(* IEC 61131-3 sources: bevling_machine/framework/sources/00_Types, 16 files *)

(* ---- E_AutoStep.st ---- *)
(* 模块说明：自动主流程步骤。正常循环从送料等料开始，切割完成后执行三路收尾。 *)
{attribute 'qualified_only'}
TYPE E_AutoStep :
(
    Idle := 0, (* 主流程待机 *)
    FeedWait := 10, (* 正常送料等料，可长期等待 *)
    StopFeed := 20, (* 撤销皮带运行并等待停止 *)
    Push := 30, (* G3 推动气缸动作 *)
    Clearance := 40, (* 并行避让 P/Q，全完成后继续 *)
    Rotate := 50, (* D8 平台旋转到配方角度 *)
    PressDown := 60, (* G1 下压到位 *)
    KnifeDown := 70, (* G9 盘刀下降到位 *)
    SpindleOn := 80, (* D3 盘刀运行状态建立 *)
    Cutting := 90, (* D2 走刀和 G6 吹气，等待指定行程到位 *)
    StopCut := 100, (* 停止盘刀和吹气 *)
    PostCut := 110, (* 抬刀、抬压、并行三路收尾 *)
    Complete := 120, (* 整循环完成，连续模式回送料 *)
    Fault := 900 (* 自动流程错误，退出执行后复位 *)
);
END_TYPE

(* ---- E_DeviceAction.st ---- *)
(* 模块说明：统一设备动作类型。未请求或停止时取消动作；定位完成依据本次命令序号判断。 *)
{attribute 'qualified_only'}
TYPE E_DeviceAction :
(
    None := 0, (* 无动作请求，取消当前动作 *)
    Position := 1, (* 定位到指定目标，等待本次序号完成 *)
    Run := 2, (* 保持连续运行请求 *)
    Jog := 3, (* 保持点动，速度正负决定方向 *)
    Stop := 4, (* 取消动作，停止运行 *)
    Home := 5 (* 回零：按轴配置的回零方式寻找原点，完成后把轴坐标设为回零坐标 *)
);
END_TYPE

(* ---- E_DeviceKind.st ---- *)
(* 模块说明：设备适配类型，由设备管理器选择轴、电机、气缸或阀的执行入口。 *)
{attribute 'qualified_only'}
TYPE E_DeviceKind :
(
    Unused := 0, (* 保留，不调度 *)
    Axis := 1, (* 定位轴 *)
    Motor := 2, (* 连续电机 *)
    Cylinder := 3, (* 两端动作气缸 *)
    Valve := 4 (* 开关阀 *)
);
END_TYPE

(* ---- E_MachineMode.st ---- *)
(* 模块说明：操作模式。手动与自动分别提出动作请求，共用设备执行和互锁。 *)
{attribute 'qualified_only'}
TYPE E_MachineMode :
(
    Manual := 0, (* 手动点动/单机构调试 *)
    Automatic := 1 (* 自动循环工序 *)
);
END_TYPE

(* ---- E_MachineState.st ---- *)
(* 模块说明：整机运行状态。停止或报警复位后须重新初始化，启动命令不会跳过初始化。 *)
{attribute 'qualified_only'}
TYPE E_MachineState :
(
    Stopped := 0, (* 停止，须初始化 *)
    Initializing := 10, (* 初始化中 *)
    Ready := 20, (* 初始化完成，等待自动启动 *)
    Manual := 30, (* 手动控制中 *)
    Automatic := 40, (* 自动工序运行中，包含正常等料 *)
    Fault := 90 (* 报警锁存，清除原因后复位 *)
);
END_TYPE

(* ---- ST_DeviceCommand.st ---- *)
(* 模块说明：上层发给单个设备的请求。定位每次换新序号；连续运行和点动期间保持请求。 *)
TYPE ST_DeviceCommand :
STRUCT
eAction : E_DeviceAction; (* 动作类型：无请求、定位、连续运行、点动或停止，见 E_DeviceAction。 *)
udiID : UDINT; (* 本次命令序号，0 无效；发起新定位时换新序号。 *)
lrTarget : LREAL; (* 目标工程位置；气缸使用约定的 0/1 端点，连续运行和点动不使用该位置。 *)
lrVelocity : LREAL; (* 请求速度，单位随设备工程单位定义；尚未完成实机标定。 *)
END_STRUCT
END_TYPE

(* ---- ST_DeviceConfig.st ---- *)
(* 模块说明：设备类型、行程范围和仿真参数。当前工程单位与时间均为仿真示例，尚未完成实机标定。 *)
TYPE ST_DeviceConfig :
STRUCT
	eKind : E_DeviceKind; (* 设备类型，决定调用哪一种设备适配功能块。 *)
	lrInitialPosition : LREAL; (* 首次进入仿真时的初始位置，不是实机回原点结果。 *)
	lrMinPosition : LREAL := -1000.0; (* 示例软行程下限，单位随机构定义。 *)
	lrMaxPosition : LREAL := 1000.0; (* 示例软行程上限，单位随机构定义。 *)
	lrMaxVelocity : LREAL := 100.0; (* 允许请求的最大速度，用于仿真命令范围检查。 *)
	tSimAction : TIME := T#500MS; (* 仿真单次定位/建立运行状态所需时间，不代表实际机械动作时间。 *)
	lrMaxAcceleration : LREAL := 50.0; (* 真实轴加速度上限，mm/s2；仿真不使用该字段。 *)
	lrMaxDeceleration : LREAL := 50.0; (* 真实轴减速度上限，mm/s2；仿真不使用该字段。 *)
	xAbsoluteAllowed : BOOL := FALSE; (* 真实轴是否允许绝对定位；未回零时必须保持 FALSE。 *)
END_STRUCT
END_TYPE

(* ---- ST_DeviceStatus.st ---- *)
(* 模块说明：单个设备的执行反馈。收到命令与完成命令是两个状态，不能只看忙标志判断完成。 *)
TYPE ST_DeviceStatus :
STRUCT
xReady : BOOL; (* 设备已使能且无故障，允许接收命令；不表示动作已经完成。 *)
xBusy : BOOL; (* 当前动作正在执行，定位完成或停止后清除。 *)
xActive : BOOL; (* 连续运行已建立或点动正在进行；定位动作完成后不保持该标志。 *)
xError : BOOL; (* 本设备或本子流程发生故障；具体原因见对应错误码。 *)
udiErrorID : UDINT; (* 错误码；0 表示无错误，设备或流程发生异常时赋值。 *)
udiAcceptedID : UDINT; (* 设备已接收的命令序号，用于区别尚未接收与正在执行。 *)
udiCompletedID : UDINT; (* 设备已完成的命令序号；应与本次 udiID 匹配后再切换步骤。 *)
lrPosition : LREAL; (* 实际或仿真反馈位置；气缸 0/1 的方向见设备编号说明。 *)
xRealActive : BOOL; (* TRUE 表示该编号当前由真实执行后端接管，不是仿真模型；默认 FALSE。 *)
xHomed : BOOL; (* 真实轴本次上电后已完成回零；仿真设备恒为 FALSE。回零成功前绝对定位会被拒绝。 *)
END_STRUCT
END_TYPE

(* ---- ST_MachineStatus.st ---- *)
(* 模块说明：提供给监控和上位机的整机状态。可从主步骤、支线步骤、报警和互锁阻挡编号定位等待原因。 *)
TYPE ST_MachineStatus :
STRUCT
	eState : E_MachineState; (* 整机状态，见 E_MachineState；调试时先确认是否已初始化及处于正确模式。 *)
	eMode : E_MachineMode; (* 本地模式旋钮的当前选择：Manual 手动，Automatic 自动；上位机仅可读取。 *)
	eAutoStep : E_AutoStep; (* 自动主流程步骤；送料、避让、切割、收尾等状态见 E_AutoStep。 *)
	xSimulation : BOOL; (* TRUE 使用内部仿真；当前 FALSE 报未实现 3001，不会接管真实运动。 *)
	xRealBackendAvailable : BOOL; (* 真实设备适配是否已具备；当前框架固定 FALSE。 *)
	xRemoteStartStopAllowed : BOOL; (* 当前是否允许上位机启停，供只读状态发布；与物理手动/自动模式独立。 *)
	xInitialized : BOOL; (* 初始化完成标志；停止、运行中切换模式或故障会清除。 *)
	xReady : BOOL; (* 整机已经初始化并处于 Ready 状态，可接受自动启动；手动状态下不置该位。 *)
	xMaterialAtLength : BOOL; (* 定长光电到位状态；自动送料须先离开再到位，并满足 D5 下降。 *)
	xCycleComplete : BOOL; (* 一个扫描周期的整循环完成脉冲，可用于计数或上位机提示。 *)
	udiCycleCount : UDINT; (* 已完成的自动整循环计数；包括机械手移料等三路收尾。 *)
	udiAlarm : UDINT; (* 整机锁存报警码；0 无报警，1001 安全许可，3001 实机未接入，10000+索引为设备故障。 *)
	uiBlockedDevice : UINT; (* 本扫描最后一个被互锁阻挡的设备索引；0 表示无阻挡，可结合设备状态排查。 *)
	uiManualReject : UINT; (* 本扫描最后一个被拒绝的手动设备索引；0 无拒绝，检查相反按钮或动作类型。 *)
	uiClearLengthStep : UINT; (* 避让支线 P 的当前步骤：10 升起 D5，20 移开 D4，1000 完成。 *)
	uiClearTransferStep : UINT; (* 避让支线 Q 当前步骤：10 降 G4，20 松 G3，30 降 G2，1000 完成。 *)
	uiPostStep : UINT; (* 收尾总步骤：10 抬刀，20 抬压，30 等待三路完成，1000 结束。 *)
	uiReturnKnifeStep : UINT; (* 收尾支线 A：10 喷油，20 D2 回刀，1000 完成。 *)
	uiUnloadStep : UINT; (* 机械手移料支线 B 步骤，10..110 每步加 10，1000 完成；详见 FB_Unload。 *)
	uiResetLengthStep : UINT; (* 收尾支线 C：10 D4 定位，20 D5 下降，30 确认下降，1000 完成。 *)
	uiInitializeStep : UINT; (* 初始化步骤：10 整理刀/压/夹爪，20 避让，25 真实轴回零，30 初始定位，40 定长下降，1000 完成。 *)
	uiActiveMaterialModel : UINT; (* 已采纳的运行料型，取自运行配方；可能与尚未生效的参数区不同。 *)
	wRemoteAckSequence : WORD; (* 整机已处理的上位机命令序号；应结合 uiRemoteResult 判断是否接受。 *)
	uiRemoteResult : UINT; (* 远程处理结果：0 接受，1 未授权，2 不支持命令，3 状态/本地停止不允许，4 验证模式禁止自动，5 配方不合法。 *)
	xAnyRealDevice : BOOL; (* 是否有任意设备由真实轴接管；TRUE 时安全源与状态发布走混跑逻辑。 *)
	xRelativeVerify : BOOL; (* 当前是否处于相对验证模式；此模式下绝对位置不作生产依据，禁止启动自动。 *)
	xSafetyBypassed : BOOL; (* 安全许可是否由两级软件旁路放行；仅调试期可为 TRUE。 *)
	uiSafetySource : UINT; (* 安全许可来源：0 仿真源，1 真实源，2 调试旁路。 *)
	wRealDeviceMask : WORD; (* 真实设备接管掩码，第 i 位置位表示设备 i 走真实轴；供上位机核对。 *)
	uiInitReject : UINT; (* 初始化被拒绝的原因：0 未拒绝；回零已并入初始化流程，当前无拒绝分支，字段预留。 *)
	xRealAxesHomed : BOOL; (* 所有已接管的真实轴都已完成回零；未接真实轴时为 TRUE。 *)
	xRunState : BOOL; (* 运行态锁存：按启动置 TRUE，按停止、安全许可丢失或进故障清 FALSE；没有它无法区分"锁存未解除"和"按钮没接"。 *)
END_STRUCT
END_TYPE

(* ---- ST_ManualCommand.st ---- *)
(* 模块说明：手动按钮接口。点动和运行按住有效，定位使用上升沿；手动请求同样经过互锁。 *)
TYPE ST_ManualCommand :
STRUCT
xJogPositive : BOOL; (* 手动正向点动，按住有效，释放后取消；只支持定位轴。 *)
xJogNegative : BOOL; (* 手动反向点动，按住有效；与正向同时按下会被拒绝。 *)
xMove : BOOL; (* 手动定位按钮，上升沿锁存目标，动作保持到本次序号完成。 *)
xHome : BOOL; (* 手动回零按钮，上升沿触发一次，动作保持到本次回零完成；只支持真实轴 D2/D8，D3 盘刀为连续旋转主轴不回零。 *)
xRun : BOOL; (* 手动连续运行按钮，按住有效、松开停止，仅支持 D1/D3/G5/G6；D3 接真实轴后由驱动器带载运行。 *)
lrTarget : LREAL; (* 目标工程位置；气缸使用约定的 0/1 端点，连续运行和点动不使用该位置。 *)
lrVelocity : LREAL := 100.0; (* 请求速度，单位随设备工程单位定义；尚未完成实机标定。 *)
END_STRUCT
END_TYPE

(* ---- ST_OperatorCommand.st ---- *)
(* 模块说明：由本地实体面板解码形成的整机命令。模式取自旋钮，初始化/启动/复位取按钮；运行态由 FB_Machine 锁存。 *)
TYPE ST_OperatorCommand :
STRUCT
eMode : E_MachineMode := E_MachineMode.Manual; (* 本地模式旋钮的当前选择：Manual 手动，Automatic 自动；上位机仅可读取。 *)
xInitialize : BOOL; (* 初始化请求，上升沿有效；只允许从停止且许可满足时进入。 *)
xStart : BOOL; (* 自动启动请求，上升沿有效；须先初始化到 Ready。 *)
xStop : BOOL; (* 停止事件，兼容保留：远程停止帧仍会写一个扫描；物理停止按钮走 xRunStop。 *)
xResetAlarm : BOOL; (* 报警复位请求，上升沿有效；原因清除后复位，不会自动重新启动。 *)
xContinuous : BOOL; (* TRUE 连续循环；FALSE 在当前完整循环结束后回到就绪。 *)
xRunStart : BOOL; (* 启动按钮标准化电平，按一下一次上升沿；FB_Machine 用它的上升沿置运行态。 *)
xRunStop : BOOL; (* 停止按钮标准化电平（常闭已取反），按一下一次上升沿；FB_Machine 用它的上升沿清运行态。 *)
END_STRUCT
END_TYPE

(* ---- ST_PanelInputs.st ---- *)
(* 模块说明：实体旋钮与按钮的逻辑输入；映射层先处理常开/常闭和极性，不在此处指定物理地址。仿真使用相同格式。 *)
TYPE ST_PanelInputs :
STRUCT
xAutoMode : BOOL; (* 模式旋钮的标准化逻辑值：TRUE 自动，FALSE 手动；不是上位机设定值。 *)
xInitialize : BOOL; (* 初始化请求，上升沿有效；只允许从停止且许可满足时进入。 *)
xStart : BOOL; (* 自动启动请求，上升沿有效；须先初始化到 Ready。 *)
xStop : BOOL; (* 停止事件，兼容保留：远程停止帧仍会写一个扫描；物理停止按钮不走这里。 *)
xResetAlarm : BOOL; (* 报警复位请求，上升沿有效；原因清除后复位，不会自动重新启动。 *)
xRunStart : BOOL; (* 启动按钮原始电平，常开、按下为 TRUE；上升沿在 FB_Machine 内锁存运行态。 *)
xRunStop : BOOL; (* 停止按钮标准化电平：常闭触点已在本层取反，按下为 TRUE；上升沿清除运行态。 *)
END_STRUCT
END_TYPE

(* ---- ST_RealDeviceSettings.st ---- *)
(* 模块说明：真实设备接管与调试旁路设置。默认接管 1、2、3、8、9、10、17 七台（现场已接线的轴与气缸），其余仍走仿真。 *)
TYPE ST_RealDeviceSettings :
STRUCT
axRealDevice : ARRAY[1..17] OF BOOL :=
    [TRUE, TRUE, TRUE, FALSE, FALSE, TRUE, FALSE, TRUE, TRUE, TRUE, FALSE, FALSE, FALSE, FALSE, FALSE, FALSE, TRUE];
    (* 逐台接管开关：TRUE = 该编号走真实硬件，FALSE = 走仿真。默认 1/2/3/6/8/9/10/17 为 TRUE。
    每次上电或完整下载都会回到这个组合；要临时关某一台，在线改位即可，但重启后恢复。
    索引对照（与 GVL_DeviceIds 的对照表完全一致，换算规则：D 编号=索引，G 编号+8=索引）：
      1=D1 送料皮带    2=D2 切割走刀    3=D3 盘刀旋转    4=D4 定长平移
      5=D5 定长升降    6=D6 定长光电    7=D7 机械手平移   8=D8 平台旋转
      9=G1 下压       10=G2 侧挡升降   11=G3 侧推       12=G4 流利条升降
      13=G5 喷油      14=G6 吹气       15=G7 机械手升降  16=G8 机械手夹爪
      17=G9 盘刀升降
    本版本只有 1、2、3、8（真实轴）、6（真实光电）与 9、10、11、17（真实气缸）已实现适配；
    其中 9（G1 下压）是左右双压板，共 4 个限位、2 路阀，设备索引仍按 1 个计；
    10（G2 侧挡）是 300/450/600 三缸一组，共 6 个限位、3 路阀，索引同样按 1 个计。
    其余编号置 TRUE 会立即报 3002，不会被静默当仿真跑。
    改本数组会让整机强制回 Stopped 并要求重新初始化，见 FB_Machine 的 wRealMask 变化检测。 *)
xRelativeVerify : BOOL; (* 相对验证模式：未回零的真实轴把 Position 解释为正向 d 再反向 d 的往返；回零成功后自动改走绝对定位。 *)
xInterlockBypass : BOOL; (* 预留：手动模式已默认不做机构互锁，本开关当前不影响判定；后续手动按需补互锁时再用。 *)
xSafetyBypass : BOOL; (* 安全许可旁路一级开关；默认 FALSE，必须与二级同时置位才生效。 *)
xSafetyBypassConfirm : BOOL; (* 安全许可旁路二级确认；默认 FALSE，防止误点单开关就旁路。 *)
xUseRealMaterial : BOOL := TRUE; (* TRUE 使用真实定长光电（设备 6）的到位信号；FALSE 继续由 FB_SimPlant 产生来料。 *)
lrVerifyDistance : LREAL := 1.0; (* 相对验证单段距离，mm；首轮建议 0.5~2.0，代码内再限幅 20。 *)
lrVerifyVelocity : LREAL := 2.0; (* 相对验证速度，mm/s；只用于未回零时的低速往返验证，不再兼作手动限速。 *)
lrVerifyAcceleration : LREAL := 50.0; (* 相对验证加速度，mm/s2。 *)
lrVerifyDeceleration : LREAL := 50.0; (* 相对验证减速度，mm/s2。 *)
tVerifyDwell : TIME := T#500MS; (* 正向到位后的停留，保证 Execute 拉低至少一个扫描以形成新上升沿。 *)
lrVerifyMeasuredByHand : LREAL; (* 人工用百分表量到的正向段实际位移，mm；用于核对轴单位标定。 *)
lrHomePosition : LREAL := 0.0; (* 预留：回零完成后的坐标由轴配置的“回零坐标”决定，MC_Homing 没有 Position 入口，本字段当前不参与下发。 *)
tHomeTimeout : TIME := T#30S; (* 单轴回零超时；超时报 2004，防止找不到原点时无限等待。 *)
lrManualVelocityMax : LREAL := 200.0; (* 手动模式速度上限，mm/s（旋转轴为每秒角度）；放在结构体末尾，避免新增字段让已有在线变量错位。 *)
END_STRUCT
END_TYPE

(* ---- ST_Recipe.st ---- *)
(* 模块说明：加工配方。初始化和自动启动时校验并复制到运行配方，避免运行中参数变化影响当前工序。 *)
TYPE ST_Recipe :
STRUCT
uiMaterialModel : UINT := 300; (* 料型选择，仅支持 300/450/600，对应 G2 三个侧挡气缸；不是位移。 *)
lrCutHome : LREAL := 100.0; (* D2 切割起点，也是回刀终点；切割终点 = 该位置 + lrCutLength。 *)
lrCutLength : LREAL := 900.0; (* D2 本次切割行程；配合 lrCutHome=100 得到终点 1000。 *)
lrCutVelocity : LREAL := 200.0; (* D2 切割进给速度，mm/s；900mm 约 5 秒走完。 *)
lrReturnVelocity : LREAL := 100.0; (* D2 回刀速度，mm/s；回刀行程长，与切割速度分开设置。 *)
lrPositionVelocity : LREAL := 10.0; (* 其余定位动作的公共请求速度，当前为仿真示例。 *)
lrBeltVelocity : LREAL := 10.0; (* D1 皮带运行速度请求，当前未换算到实际驱动器单位。 *)
lrSpindleVelocity : LREAL := 50.0; (* D3 盘刀运行速度请求，mm/s；不是已标定的实际转速。自动切割默认 50。 *)
lrLengthPosition : LREAL := 100.0; (* D4 定长检测工作位置；到位后再令 D5 下降。 *)
lrLengthClear : LREAL := 0.0; (* D4 切割前避让位置；移动前须 D5 升起。 *)
lrRotateAngle : LREAL := 30; (* D8 平台旋转目标角度，示例范围为正负 360，实机角度单位待标定。 *)
lrGripperFront : LREAL := 100.0; (* D7 机械手前进取料位置。 *)
lrGripperPull : LREAL := 200.0; (* D7 夹紧后拉料目标位置。 *)
lrGripperBack : LREAL := 50.0; (* D7 松开后的抬升后退位置；到位后先下降，再最终回位。 *)
lrGripperHome : LREAL := 0.0; (* D7 机械手下降后最终回位的位置。 *)
tSpray : TIME := T#300MS; (* 收尾支线 A 的喷油保持时间；该步结束后撤销喷油请求。 *)
tStepTimeout : TIME := T#30S; (* 单动作步骤超时时间；正常送料等料阶段不套用此超时。 *)
tCutTimeout : TIME := T#30S; (* D2 切割步专用超时，独立于 tStepTimeout；加在结构体末尾，避免新增字段让已有在线变量错位。 *)
END_STRUCT
END_TYPE

(* ---- ST_RemoteCommand.st ---- *)
(* 模块说明：上位机可选启停请求，不含模式、初始化、复位或连续选择字段。参数通过独立配方接口下发。 *)
TYPE ST_RemoteCommand :
STRUCT
xStart : BOOL; (* 自动启动请求，上升沿有效；须先初始化到 Ready。 *)
xStop : BOOL; (* 普通停止，TRUE 持续有效；取消动作并清除初始化，不能替代硬件急停。 *)
END_STRUCT
END_TYPE

(* ---- ST_SimulationSettings.st ---- *)
(* 模块说明：软件仿真输入和异常注入。设备索引为 1..17，与 GVL_DeviceIds 一致。 *)
TYPE ST_SimulationSettings :
STRUCT
xSafetyOK : BOOL := TRUE; (* 安全许可接口或仿真许可，TRUE 允许；不等同于安全级急停回路。 *)
xAutoMaterial : BOOL := TRUE; (* TRUE 由仿真模型自动产生到位；FALSE 使用人工料到位输入。 *)
xMaterialSensor : BOOL; (* 手动模拟的光电到位信号，仅在 xAutoMaterial=FALSE 时使用。 *)
tMaterialDelay : TIME := T#1S; (* 满足皮带运行及定长下降条件后，仿真来料的延时时间。 *)
axStall : ARRAY[1..17] OF BOOL; (* 设备卡住注入，索引 1..17；保持忙且不完成，用于观察等待/超时。 *)
axFault : ARRAY[1..17] OF BOOL; (* 设备故障注入，索引 1..17；先清除注入，再执行报警复位。 *)
END_STRUCT
END_TYPE
